FUNCTION FC 1 : VOID
BEGIN
NETWORK
      U E 0.0
END_FUNCTION
